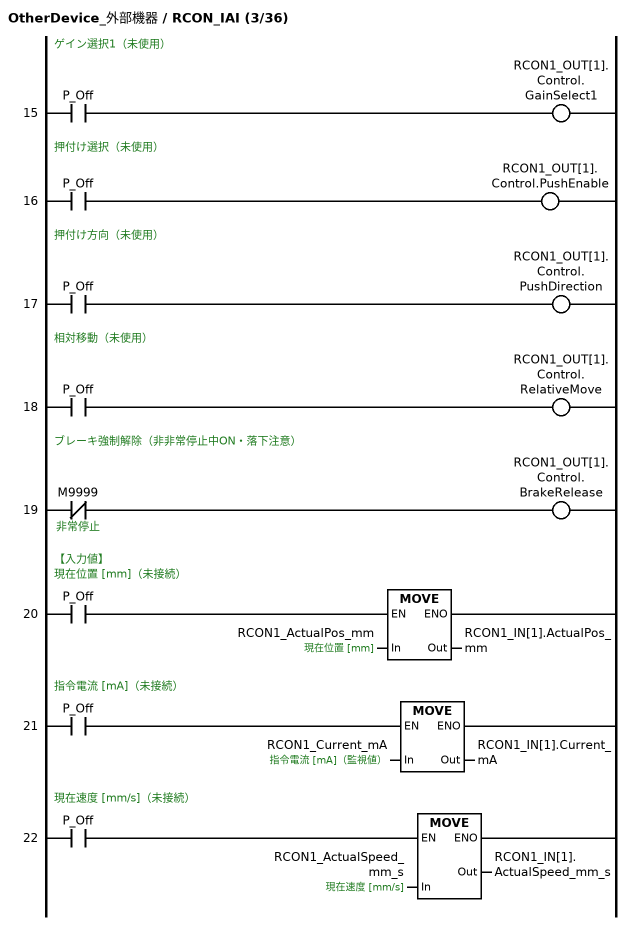
(* [picture p48: OtherDevice_外部機器 / RCON_IAI, rungs 15-22] *)
(* Rung 15: ゲイン選択1（未使用） *)
RCON1_OUT[1].Control.GainSelect1 := P_Off;
(* Rung 16: 押付け選択（未使用） *)
RCON1_OUT[1].Control.PushEnable := P_Off;
(* Rung 17: 押付け方向（未使用） *)
RCON1_OUT[1].Control.PushDirection := P_Off;
(* Rung 18: 相対移動（未使用） *)
RCON1_OUT[1].Control.RelativeMove := P_Off;
(* Rung 19: ブレーキ強制解除（非非常停止中ON・落下注意） *)
RCON1_OUT[1].Control.BrakeRelease := NOT M9999;
(* Rung 20: 【入力値】 / 現在位置 [mm]（未接続） *)
IF P_Off THEN RCON1_IN[1].ActualPos_mm := RCON1_ActualPos_mm; END_IF;
(* Rung 21: 指令電流 [mA]（未接続） *)
IF P_Off THEN RCON1_IN[1].Current_mA := RCON1_Current_mA; END_IF;
(* Rung 22: 現在速度 [mm/s]（未接続） *)
IF P_Off THEN RCON1_IN[1].ActualSpeed_mm_s := RCON1_ActualSpeed_mm_s; END_IF;

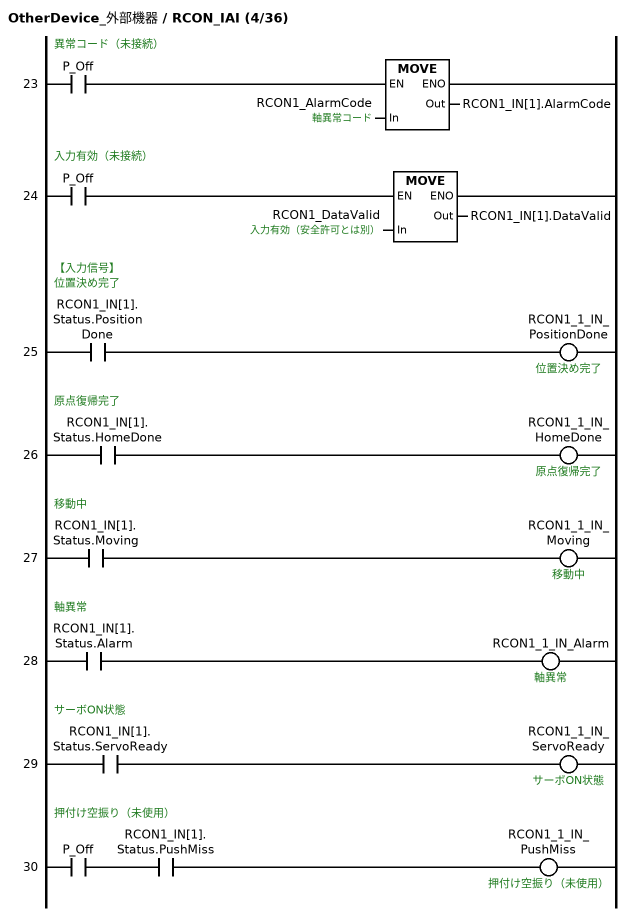
(* Rung 23: 異常コード（未接続） *)
IF P_Off THEN RCON1_IN[1].AlarmCode := RCON1_AlarmCode; END_IF;
(* Rung 24: 入力有効（未接続） *)
IF P_Off THEN RCON1_IN[1].DataValid := RCON1_DataValid; END_IF;
(* Rung 25: 【入力信号】 / 位置決め完了 *)
RCON1_1_IN_PositionDone := RCON1_IN[1].Status.PositionDone;
(* Rung 26: 原点復帰完了 *)
RCON1_1_IN_HomeDone := RCON1_IN[1].Status.HomeDone;
(* Rung 27: 移動中 *)
RCON1_1_IN_Moving := RCON1_IN[1].Status.Moving;
(* Rung 28: 軸異常 *)
RCON1_1_IN_Alarm := RCON1_IN[1].Status.Alarm;
(* Rung 29: サーボON状態 *)
RCON1_1_IN_ServoReady := RCON1_IN[1].Status.ServoReady;
(* Rung 30: 押付け空振り（未使用） *)
RCON1_1_IN_PushMiss := P_Off AND RCON1_IN[1].Status.PushMiss;

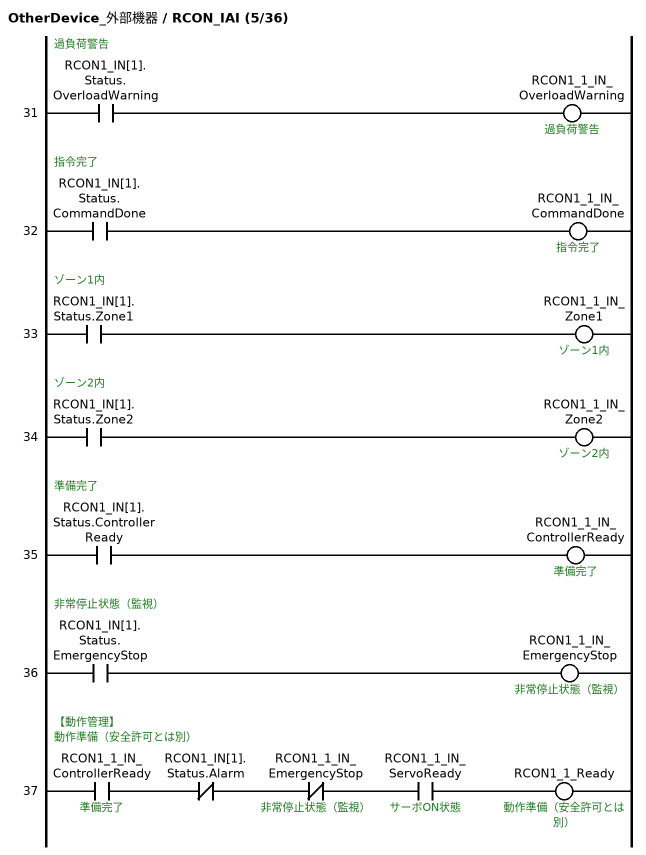
(* Rung 31: 過負荷警告 *)
RCON1_1_IN_OverloadWarning := RCON1_IN[1].Status.OverloadWarning;
(* Rung 32: 指令完了 *)
RCON1_1_IN_CommandDone := RCON1_IN[1].Status.CommandDone;
(* Rung 33: ゾーン1内 *)
RCON1_1_IN_Zone1 := RCON1_IN[1].Status.Zone1;
(* Rung 34: ゾーン2内 *)
RCON1_1_IN_Zone2 := RCON1_IN[1].Status.Zone2;
(* Rung 35: 準備完了 *)
RCON1_1_IN_ControllerReady := RCON1_IN[1].Status.ControllerReady;
(* Rung 36: 非常停止状態（監視） *)
RCON1_1_IN_EmergencyStop := RCON1_IN[1].Status.EmergencyStop;
(* Rung 37: 【動作管理】 / 動作準備（安全許可とは別） *)
RCON1_1_Ready := RCON1_1_IN_ControllerReady AND NOT RCON1_IN[1].Status.Alarm AND NOT RCON1_1_IN_EmergencyStop AND RCON1_1_IN_ServoReady;

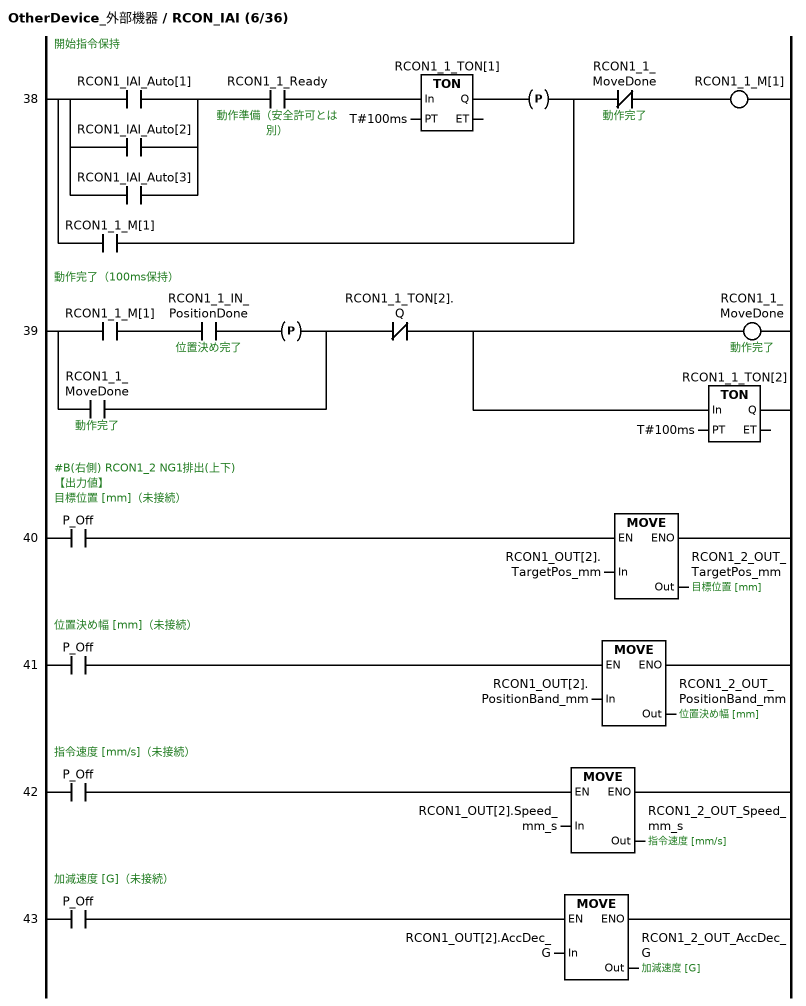
(* Rung 38: 開始指令保持 *)
RCON1_1_TON[1](In := (RCON1_IAI_Auto[1] OR RCON1_IAI_Auto[2] OR RCON1_IAI_Auto[3]) AND RCON1_1_Ready, PT := T#100ms);
_e2(CLK := RCON1_1_TON[1].Q);
RCON1_1_M[1] := (_e2.Q OR RCON1_1_M[1]) AND NOT RCON1_1_MoveDone;
(* Rung 39: 動作完了（100ms保持） *)
_e3(CLK := RCON1_1_M[1] AND RCON1_1_IN_PositionDone);
_p4 := (_e3.Q OR RCON1_1_MoveDone) AND NOT RCON1_1_TON[2].Q;
RCON1_1_MoveDone := _p4;
RCON1_1_TON[2](In := _p4, PT := T#100ms);
(* Rung 40: #B(右側) RCON1_2 NG1排出(上下) / 【出力値】 / 目標位置 [mm]（未接続） *)
IF P_Off THEN RCON1_2_OUT_TargetPos_mm := RCON1_OUT[2].TargetPos_mm; END_IF;
(* Rung 41: 位置決め幅 [mm]（未接続） *)
IF P_Off THEN RCON1_2_OUT_PositionBand_mm := RCON1_OUT[2].PositionBand_mm; END_IF;
(* Rung 42: 指令速度 [mm/s]（未接続） *)
IF P_Off THEN RCON1_2_OUT_Speed_mm_s := RCON1_OUT[2].Speed_mm_s; END_IF;
(* Rung 43: 加減速度 [G]（未接続） *)
IF P_Off THEN RCON1_2_OUT_AccDec_G := RCON1_OUT[2].AccDec_G; END_IF;

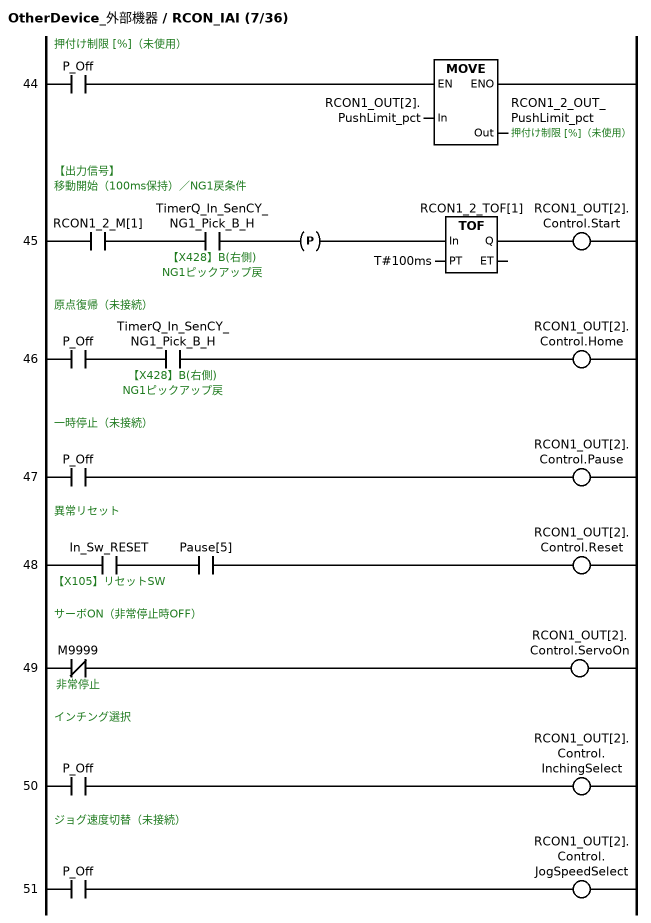
(* Rung 44: 押付け制限 [%]（未使用） *)
IF P_Off THEN RCON1_2_OUT_PushLimit_pct := RCON1_OUT[2].PushLimit_pct; END_IF;
(* Rung 45: 【出力信号】 / 移動開始（100ms保持）／NG1戻条件 *)
_e5(CLK := RCON1_2_M[1] AND TimerQ_In_SenCY_NG1_Pick_B_H);
RCON1_2_TOF[1](In := _e5.Q, PT := T#100ms);
RCON1_OUT[2].Control.Start := RCON1_2_TOF[1].Q;
(* Rung 46: 原点復帰（未接続） *)
RCON1_OUT[2].Control.Home := P_Off AND TimerQ_In_SenCY_NG1_Pick_B_H;
(* Rung 47: 一時停止（未接続） *)
RCON1_OUT[2].Control.Pause := P_Off;
(* Rung 48: 異常リセット *)
RCON1_OUT[2].Control.Reset := In_Sw_RESET AND Pause[5];
(* Rung 49: サーボON（非常停止時OFF） *)
RCON1_OUT[2].Control.ServoOn := NOT M9999;
(* Rung 50: インチング選択 *)
RCON1_OUT[2].Control.InchingSelect := P_Off;
(* Rung 51: ジョグ速度切替（未接続） *)
RCON1_OUT[2].Control.JogSpeedSelect := P_Off;

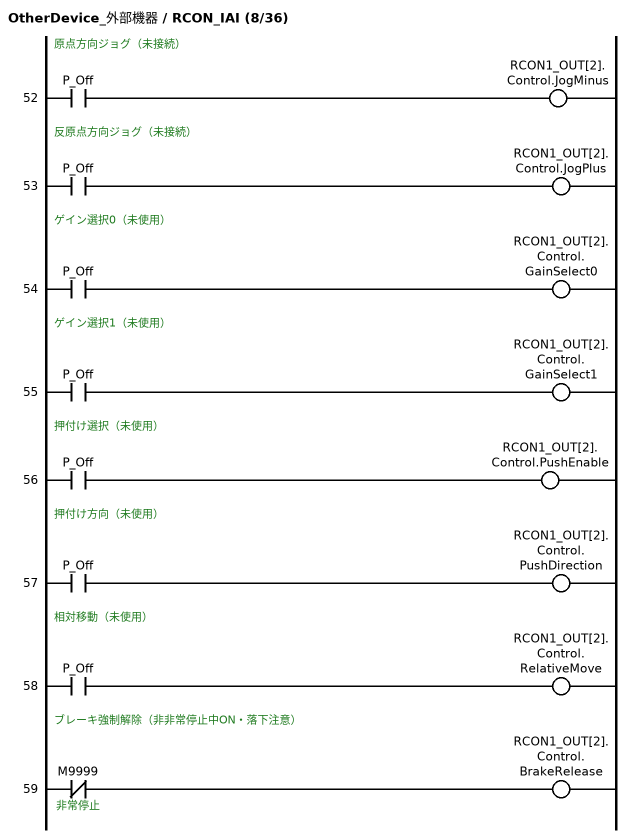
(* Rung 52: 原点方向ジョグ（未接続） *)
RCON1_OUT[2].Control.JogMinus := P_Off;
(* Rung 53: 反原点方向ジョグ（未接続） *)
RCON1_OUT[2].Control.JogPlus := P_Off;
(* Rung 54: ゲイン選択0（未使用） *)
RCON1_OUT[2].Control.GainSelect0 := P_Off;
(* Rung 55: ゲイン選択1（未使用） *)
RCON1_OUT[2].Control.GainSelect1 := P_Off;
(* Rung 56: 押付け選択（未使用） *)
RCON1_OUT[2].Control.PushEnable := P_Off;
(* Rung 57: 押付け方向（未使用） *)
RCON1_OUT[2].Control.PushDirection := P_Off;
(* Rung 58: 相対移動（未使用） *)
RCON1_OUT[2].Control.RelativeMove := P_Off;
(* Rung 59: ブレーキ強制解除（非非常停止中ON・落下注意） *)
RCON1_OUT[2].Control.BrakeRelease := NOT M9999;

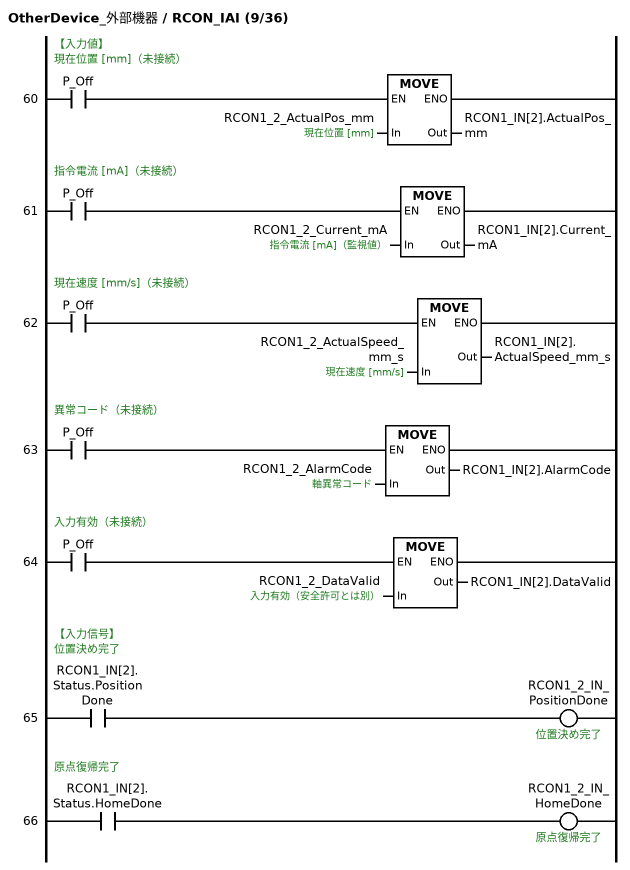
(* Rung 60: 【入力値】 / 現在位置 [mm]（未接続） *)
IF P_Off THEN RCON1_IN[2].ActualPos_mm := RCON1_2_ActualPos_mm; END_IF;
(* Rung 61: 指令電流 [mA]（未接続） *)
IF P_Off THEN RCON1_IN[2].Current_mA := RCON1_2_Current_mA; END_IF;
(* Rung 62: 現在速度 [mm/s]（未接続） *)
IF P_Off THEN RCON1_IN[2].ActualSpeed_mm_s := RCON1_2_ActualSpeed_mm_s; END_IF;
(* Rung 63: 異常コード（未接続） *)
IF P_Off THEN RCON1_IN[2].AlarmCode := RCON1_2_AlarmCode; END_IF;
(* Rung 64: 入力有効（未接続） *)
IF P_Off THEN RCON1_IN[2].DataValid := RCON1_2_DataValid; END_IF;
(* Rung 65: 【入力信号】 / 位置決め完了 *)
RCON1_2_IN_PositionDone := RCON1_IN[2].Status.PositionDone;
(* Rung 66: 原点復帰完了 *)
RCON1_2_IN_HomeDone := RCON1_IN[2].Status.HomeDone;

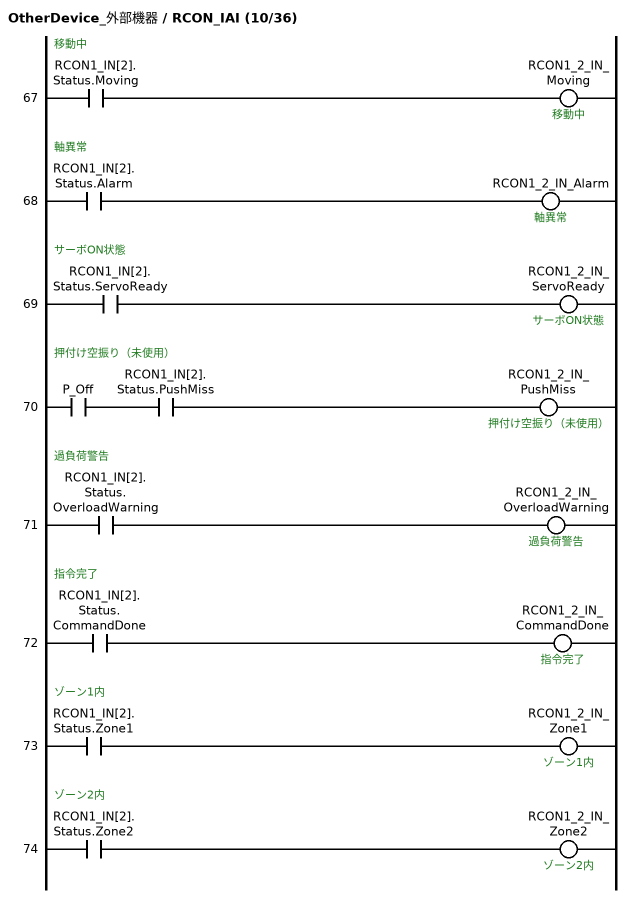
(* Rung 67: 移動中 *)
RCON1_2_IN_Moving := RCON1_IN[2].Status.Moving;
(* Rung 68: 軸異常 *)
RCON1_2_IN_Alarm := RCON1_IN[2].Status.Alarm;
(* Rung 69: サーボON状態 *)
RCON1_2_IN_ServoReady := RCON1_IN[2].Status.ServoReady;
(* Rung 70: 押付け空振り（未使用） *)
RCON1_2_IN_PushMiss := P_Off AND RCON1_IN[2].Status.PushMiss;
(* Rung 71: 過負荷警告 *)
RCON1_2_IN_OverloadWarning := RCON1_IN[2].Status.OverloadWarning;
(* Rung 72: 指令完了 *)
RCON1_2_IN_CommandDone := RCON1_IN[2].Status.CommandDone;
(* Rung 73: ゾーン1内 *)
RCON1_2_IN_Zone1 := RCON1_IN[2].Status.Zone1;
(* Rung 74: ゾーン2内 *)
RCON1_2_IN_Zone2 := RCON1_IN[2].Status.Zone2;

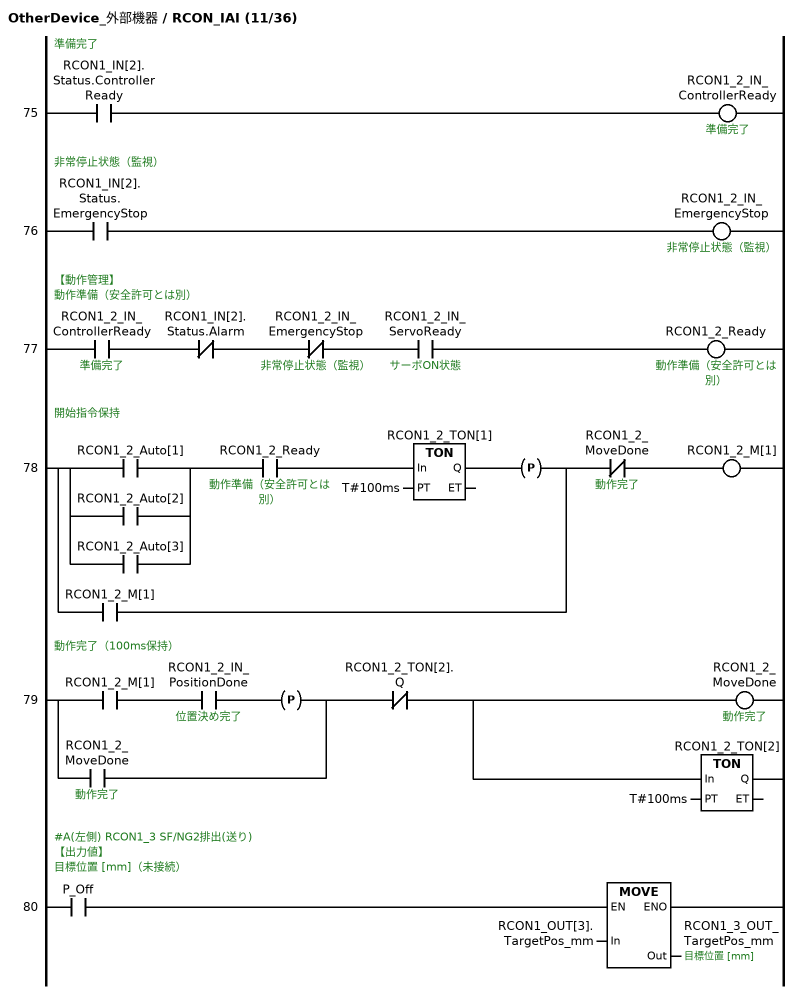
(* Rung 75: 準備完了 *)
RCON1_2_IN_ControllerReady := RCON1_IN[2].Status.ControllerReady;
(* Rung 76: 非常停止状態（監視） *)
RCON1_2_IN_EmergencyStop := RCON1_IN[2].Status.EmergencyStop;
(* Rung 77: 【動作管理】 / 動作準備（安全許可とは別） *)
RCON1_2_Ready := RCON1_2_IN_ControllerReady AND NOT RCON1_IN[2].Status.Alarm AND NOT RCON1_2_IN_EmergencyStop AND RCON1_2_IN_ServoReady;
(* Rung 78: 開始指令保持 *)
RCON1_2_TON[1](In := (RCON1_2_Auto[1] OR RCON1_2_Auto[2] OR RCON1_2_Auto[3]) AND RCON1_2_Ready, PT := T#100ms);
_e6(CLK := RCON1_2_TON[1].Q);
RCON1_2_M[1] := (_e6.Q OR RCON1_2_M[1]) AND NOT RCON1_2_MoveDone;
(* Rung 79: 動作完了（100ms保持） *)
_e7(CLK := RCON1_2_M[1] AND RCON1_2_IN_PositionDone);
_p8 := (_e7.Q OR RCON1_2_MoveDone) AND NOT RCON1_2_TON[2].Q;
RCON1_2_MoveDone := _p8;
RCON1_2_TON[2](In := _p8, PT := T#100ms);
(* Rung 80: #A(左側) RCON1_3 SF/NG2排出(送り) / 【出力値】 / 目標位置 [mm]（未接続） *)
IF P_Off THEN RCON1_3_OUT_TargetPos_mm := RCON1_OUT[3].TargetPos_mm; END_IF;

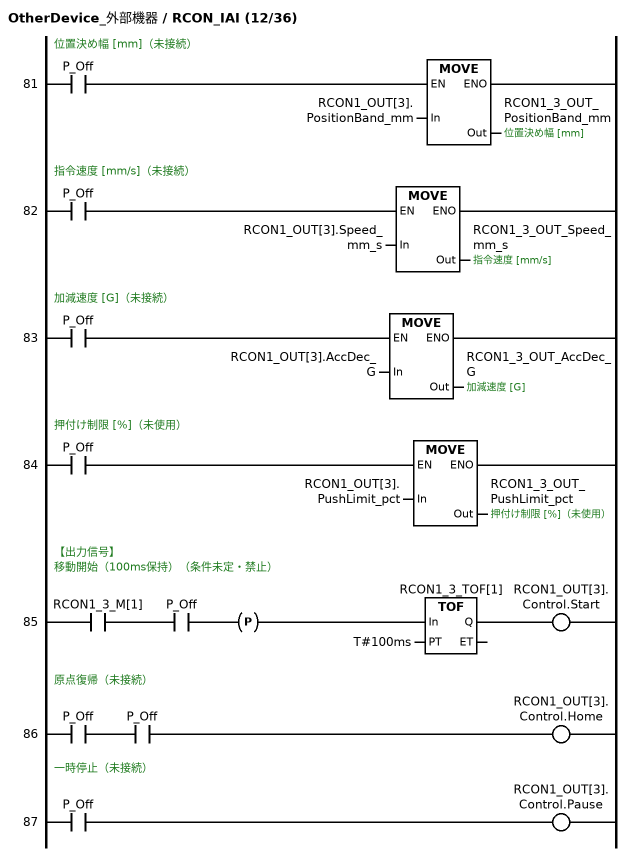
(* Rung 81: 位置決め幅 [mm]（未接続） *)
IF P_Off THEN RCON1_3_OUT_PositionBand_mm := RCON1_OUT[3].PositionBand_mm; END_IF;
(* Rung 82: 指令速度 [mm/s]（未接続） *)
IF P_Off THEN RCON1_3_OUT_Speed_mm_s := RCON1_OUT[3].Speed_mm_s; END_IF;
(* Rung 83: 加減速度 [G]（未接続） *)
IF P_Off THEN RCON1_3_OUT_AccDec_G := RCON1_OUT[3].AccDec_G; END_IF;
(* Rung 84: 押付け制限 [%]（未使用） *)
IF P_Off THEN RCON1_3_OUT_PushLimit_pct := RCON1_OUT[3].PushLimit_pct; END_IF;
(* Rung 85: 【出力信号】 / 移動開始（100ms保持）（条件未定・禁止） *)
_e9(CLK := RCON1_3_M[1] AND P_Off);
RCON1_3_TOF[1](In := _e9.Q, PT := T#100ms);
RCON1_OUT[3].Control.Start := RCON1_3_TOF[1].Q;
(* Rung 86: 原点復帰（未接続） *)
RCON1_OUT[3].Control.Home := P_Off AND P_Off;
(* Rung 87: 一時停止（未接続） *)
RCON1_OUT[3].Control.Pause := P_Off;

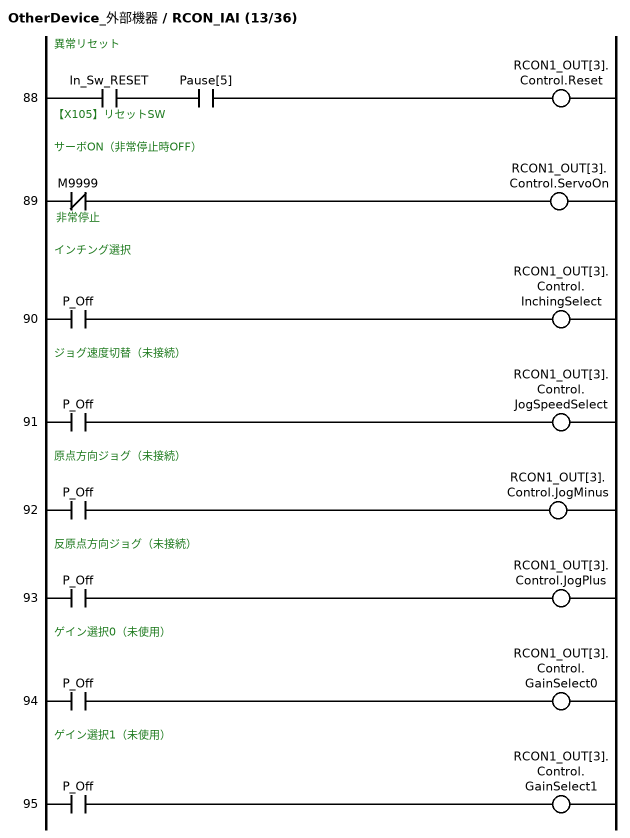
(* Rung 88: 異常リセット *)
RCON1_OUT[3].Control.Reset := In_Sw_RESET AND Pause[5];
(* Rung 89: サーボON（非常停止時OFF） *)
RCON1_OUT[3].Control.ServoOn := NOT M9999;
(* Rung 90: インチング選択 *)
RCON1_OUT[3].Control.InchingSelect := P_Off;
(* Rung 91: ジョグ速度切替（未接続） *)
RCON1_OUT[3].Control.JogSpeedSelect := P_Off;
(* Rung 92: 原点方向ジョグ（未接続） *)
RCON1_OUT[3].Control.JogMinus := P_Off;
(* Rung 93: 反原点方向ジョグ（未接続） *)
RCON1_OUT[3].Control.JogPlus := P_Off;
(* Rung 94: ゲイン選択0（未使用） *)
RCON1_OUT[3].Control.GainSelect0 := P_Off;
(* Rung 95: ゲイン選択1（未使用） *)
RCON1_OUT[3].Control.GainSelect1 := P_Off;

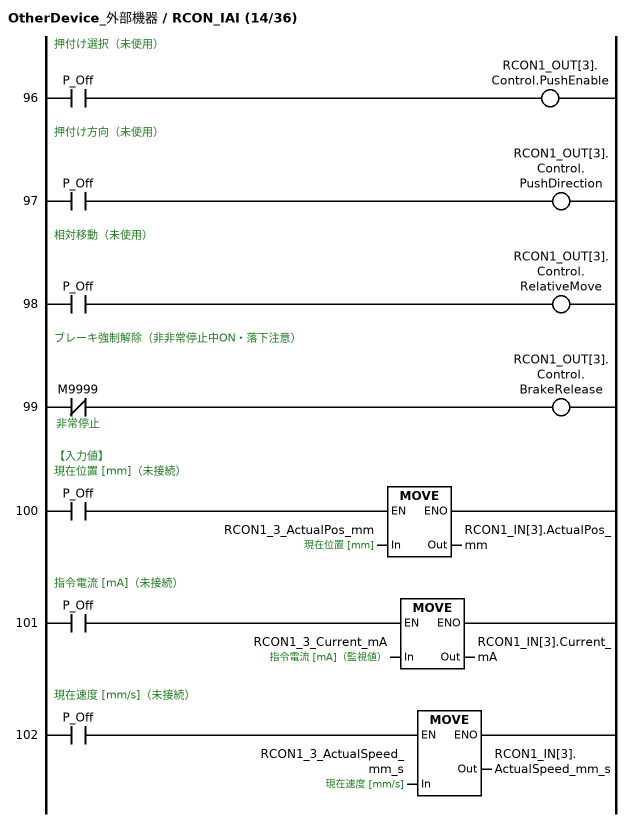
(* Rung 96: 押付け選択（未使用） *)
RCON1_OUT[3].Control.PushEnable := P_Off;
(* Rung 97: 押付け方向（未使用） *)
RCON1_OUT[3].Control.PushDirection := P_Off;
(* Rung 98: 相対移動（未使用） *)
RCON1_OUT[3].Control.RelativeMove := P_Off;
(* Rung 99: ブレーキ強制解除（非非常停止中ON・落下注意） *)
RCON1_OUT[3].Control.BrakeRelease := NOT M9999;
(* Rung 100: 【入力値】 / 現在位置 [mm]（未接続） *)
IF P_Off THEN RCON1_IN[3].ActualPos_mm := RCON1_3_ActualPos_mm; END_IF;
(* Rung 101: 指令電流 [mA]（未接続） *)
IF P_Off THEN RCON1_IN[3].Current_mA := RCON1_3_Current_mA; END_IF;
(* Rung 102: 現在速度 [mm/s]（未接続） *)
IF P_Off THEN RCON1_IN[3].ActualSpeed_mm_s := RCON1_3_ActualSpeed_mm_s; END_IF;

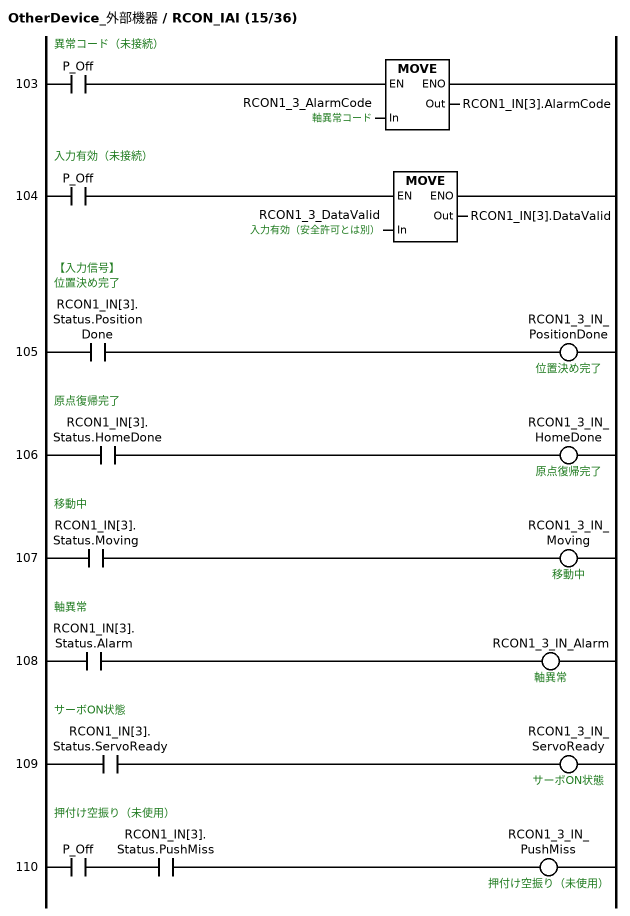
(* Rung 103: 異常コード（未接続） *)
IF P_Off THEN RCON1_IN[3].AlarmCode := RCON1_3_AlarmCode; END_IF;
(* Rung 104: 入力有効（未接続） *)
IF P_Off THEN RCON1_IN[3].DataValid := RCON1_3_DataValid; END_IF;
(* Rung 105: 【入力信号】 / 位置決め完了 *)
RCON1_3_IN_PositionDone := RCON1_IN[3].Status.PositionDone;
(* Rung 106: 原点復帰完了 *)
RCON1_3_IN_HomeDone := RCON1_IN[3].Status.HomeDone;
(* Rung 107: 移動中 *)
RCON1_3_IN_Moving := RCON1_IN[3].Status.Moving;
(* Rung 108: 軸異常 *)
RCON1_3_IN_Alarm := RCON1_IN[3].Status.Alarm;
(* Rung 109: サーボON状態 *)
RCON1_3_IN_ServoReady := RCON1_IN[3].Status.ServoReady;
(* Rung 110: 押付け空振り（未使用） *)
RCON1_3_IN_PushMiss := P_Off AND RCON1_IN[3].Status.PushMiss;

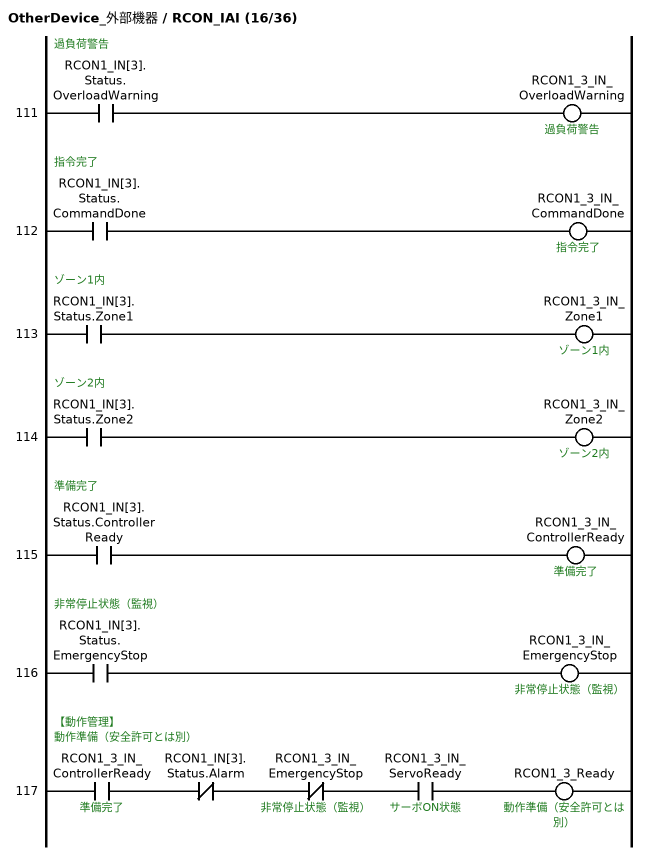
(* Rung 111: 過負荷警告 *)
RCON1_3_IN_OverloadWarning := RCON1_IN[3].Status.OverloadWarning;
(* Rung 112: 指令完了 *)
RCON1_3_IN_CommandDone := RCON1_IN[3].Status.CommandDone;
(* Rung 113: ゾーン1内 *)
RCON1_3_IN_Zone1 := RCON1_IN[3].Status.Zone1;
(* Rung 114: ゾーン2内 *)
RCON1_3_IN_Zone2 := RCON1_IN[3].Status.Zone2;
(* Rung 115: 準備完了 *)
RCON1_3_IN_ControllerReady := RCON1_IN[3].Status.ControllerReady;
(* Rung 116: 非常停止状態（監視） *)
RCON1_3_IN_EmergencyStop := RCON1_IN[3].Status.EmergencyStop;
(* Rung 117: 【動作管理】 / 動作準備（安全許可とは別） *)
RCON1_3_Ready := RCON1_3_IN_ControllerReady AND NOT RCON1_IN[3].Status.Alarm AND NOT RCON1_3_IN_EmergencyStop AND RCON1_3_IN_ServoReady;

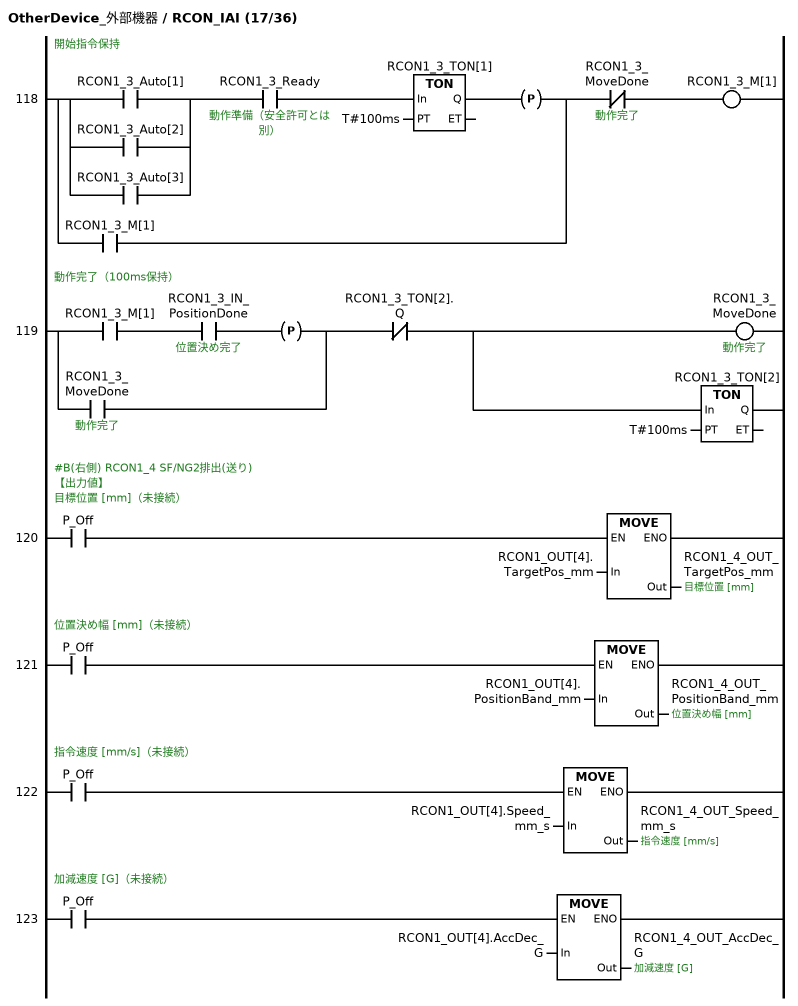
(* Rung 118: 開始指令保持 *)
RCON1_3_TON[1](In := (RCON1_3_Auto[1] OR RCON1_3_Auto[2] OR RCON1_3_Auto[3]) AND RCON1_3_Ready, PT := T#100ms);
_e10(CLK := RCON1_3_TON[1].Q);
RCON1_3_M[1] := (_e10.Q OR RCON1_3_M[1]) AND NOT RCON1_3_MoveDone;
(* Rung 119: 動作完了（100ms保持） *)
_e11(CLK := RCON1_3_M[1] AND RCON1_3_IN_PositionDone);
_p12 := (_e11.Q OR RCON1_3_MoveDone) AND NOT RCON1_3_TON[2].Q;
RCON1_3_MoveDone := _p12;
RCON1_3_TON[2](In := _p12, PT := T#100ms);
(* Rung 120: #B(右側) RCON1_4 SF/NG2排出(送り) / 【出力値】 / 目標位置 [mm]（未接続） *)
IF P_Off THEN RCON1_4_OUT_TargetPos_mm := RCON1_OUT[4].TargetPos_mm; END_IF;
(* Rung 121: 位置決め幅 [mm]（未接続） *)
IF P_Off THEN RCON1_4_OUT_PositionBand_mm := RCON1_OUT[4].PositionBand_mm; END_IF;
(* Rung 122: 指令速度 [mm/s]（未接続） *)
IF P_Off THEN RCON1_4_OUT_Speed_mm_s := RCON1_OUT[4].Speed_mm_s; END_IF;
(* Rung 123: 加減速度 [G]（未接続） *)
IF P_Off THEN RCON1_4_OUT_AccDec_G := RCON1_OUT[4].AccDec_G; END_IF;

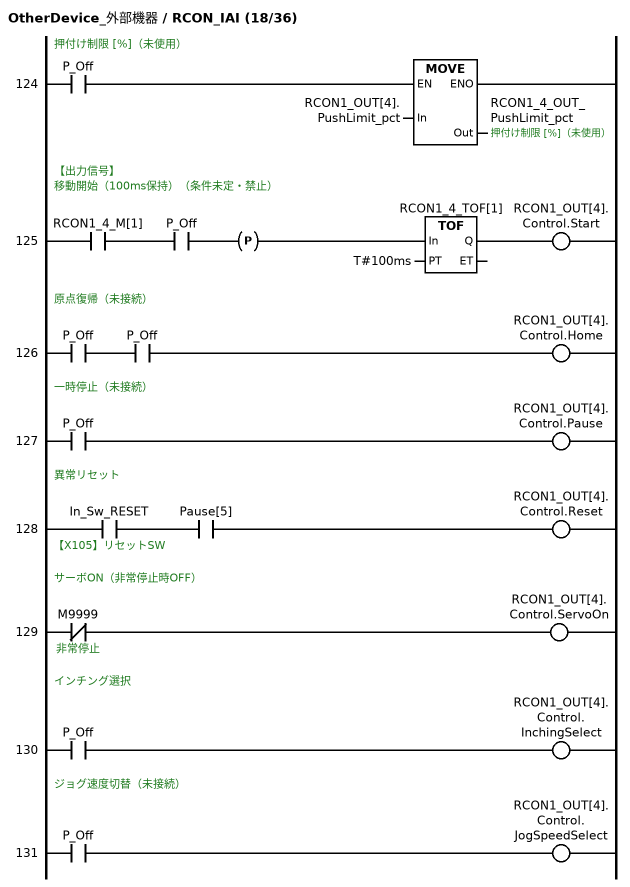
(* Rung 124: 押付け制限 [%]（未使用） *)
IF P_Off THEN RCON1_4_OUT_PushLimit_pct := RCON1_OUT[4].PushLimit_pct; END_IF;
(* Rung 125: 【出力信号】 / 移動開始（100ms保持）（条件未定・禁止） *)
_e13(CLK := RCON1_4_M[1] AND P_Off);
RCON1_4_TOF[1](In := _e13.Q, PT := T#100ms);
RCON1_OUT[4].Control.Start := RCON1_4_TOF[1].Q;
(* Rung 126: 原点復帰（未接続） *)
RCON1_OUT[4].Control.Home := P_Off AND P_Off;
(* Rung 127: 一時停止（未接続） *)
RCON1_OUT[4].Control.Pause := P_Off;
(* Rung 128: 異常リセット *)
RCON1_OUT[4].Control.Reset := In_Sw_RESET AND Pause[5];
(* Rung 129: サーボON（非常停止時OFF） *)
RCON1_OUT[4].Control.ServoOn := NOT M9999;
(* Rung 130: インチング選択 *)
RCON1_OUT[4].Control.InchingSelect := P_Off;
(* Rung 131: ジョグ速度切替（未接続） *)
RCON1_OUT[4].Control.JogSpeedSelect := P_Off;

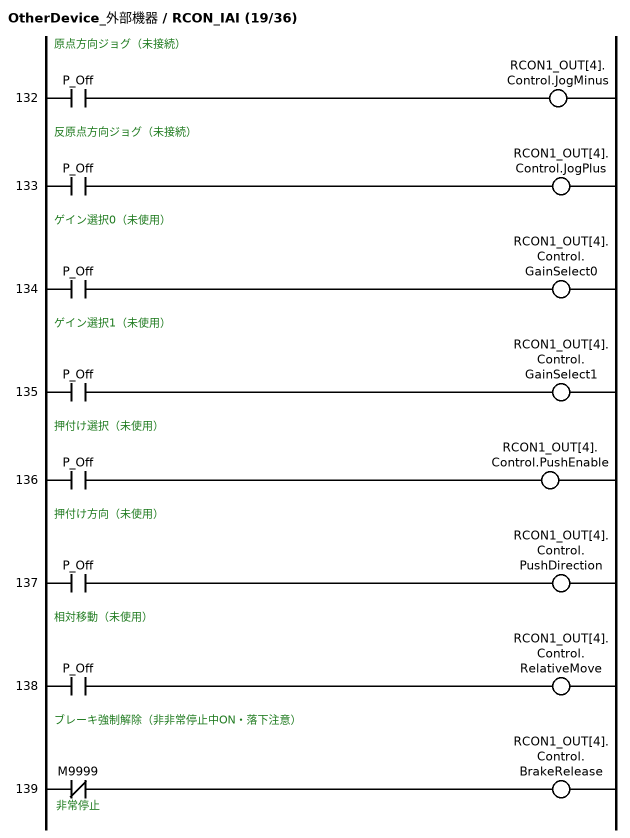
(* Rung 132: 原点方向ジョグ（未接続） *)
RCON1_OUT[4].Control.JogMinus := P_Off;
(* Rung 133: 反原点方向ジョグ（未接続） *)
RCON1_OUT[4].Control.JogPlus := P_Off;
(* Rung 134: ゲイン選択0（未使用） *)
RCON1_OUT[4].Control.GainSelect0 := P_Off;
(* Rung 135: ゲイン選択1（未使用） *)
RCON1_OUT[4].Control.GainSelect1 := P_Off;
(* Rung 136: 押付け選択（未使用） *)
RCON1_OUT[4].Control.PushEnable := P_Off;
(* Rung 137: 押付け方向（未使用） *)
RCON1_OUT[4].Control.PushDirection := P_Off;
(* Rung 138: 相対移動（未使用） *)
RCON1_OUT[4].Control.RelativeMove := P_Off;
(* Rung 139: ブレーキ強制解除（非非常停止中ON・落下注意） *)
RCON1_OUT[4].Control.BrakeRelease := NOT M9999;

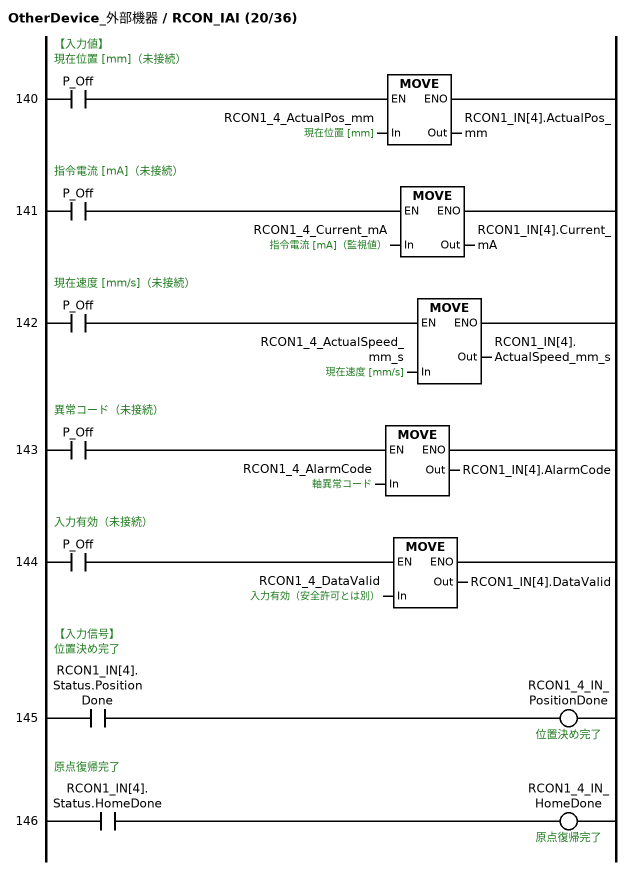
(* Rung 140: 【入力値】 / 現在位置 [mm]（未接続） *)
IF P_Off THEN RCON1_IN[4].ActualPos_mm := RCON1_4_ActualPos_mm; END_IF;
(* Rung 141: 指令電流 [mA]（未接続） *)
IF P_Off THEN RCON1_IN[4].Current_mA := RCON1_4_Current_mA; END_IF;
(* Rung 142: 現在速度 [mm/s]（未接続） *)
IF P_Off THEN RCON1_IN[4].ActualSpeed_mm_s := RCON1_4_ActualSpeed_mm_s; END_IF;
(* Rung 143: 異常コード（未接続） *)
IF P_Off THEN RCON1_IN[4].AlarmCode := RCON1_4_AlarmCode; END_IF;
(* Rung 144: 入力有効（未接続） *)
IF P_Off THEN RCON1_IN[4].DataValid := RCON1_4_DataValid; END_IF;
(* Rung 145: 【入力信号】 / 位置決め完了 *)
RCON1_4_IN_PositionDone := RCON1_IN[4].Status.PositionDone;
(* Rung 146: 原点復帰完了 *)
RCON1_4_IN_HomeDone := RCON1_IN[4].Status.HomeDone;

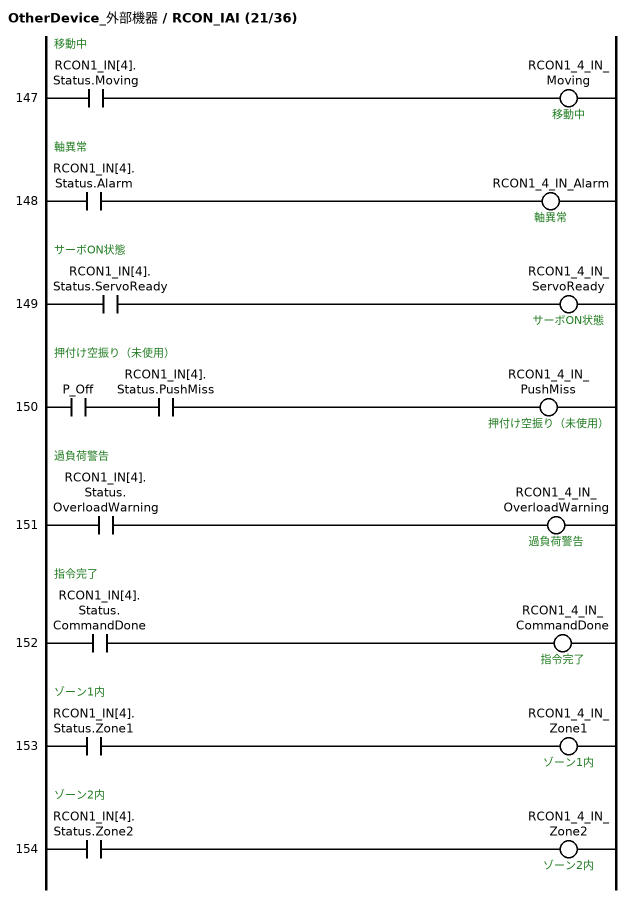
(* Rung 147: 移動中 *)
RCON1_4_IN_Moving := RCON1_IN[4].Status.Moving;
(* Rung 148: 軸異常 *)
RCON1_4_IN_Alarm := RCON1_IN[4].Status.Alarm;
(* Rung 149: サーボON状態 *)
RCON1_4_IN_ServoReady := RCON1_IN[4].Status.ServoReady;
(* Rung 150: 押付け空振り（未使用） *)
RCON1_4_IN_PushMiss := P_Off AND RCON1_IN[4].Status.PushMiss;
(* Rung 151: 過負荷警告 *)
RCON1_4_IN_OverloadWarning := RCON1_IN[4].Status.OverloadWarning;
(* Rung 152: 指令完了 *)
RCON1_4_IN_CommandDone := RCON1_IN[4].Status.CommandDone;
(* Rung 153: ゾーン1内 *)
RCON1_4_IN_Zone1 := RCON1_IN[4].Status.Zone1;
(* Rung 154: ゾーン2内 *)
RCON1_4_IN_Zone2 := RCON1_IN[4].Status.Zone2;

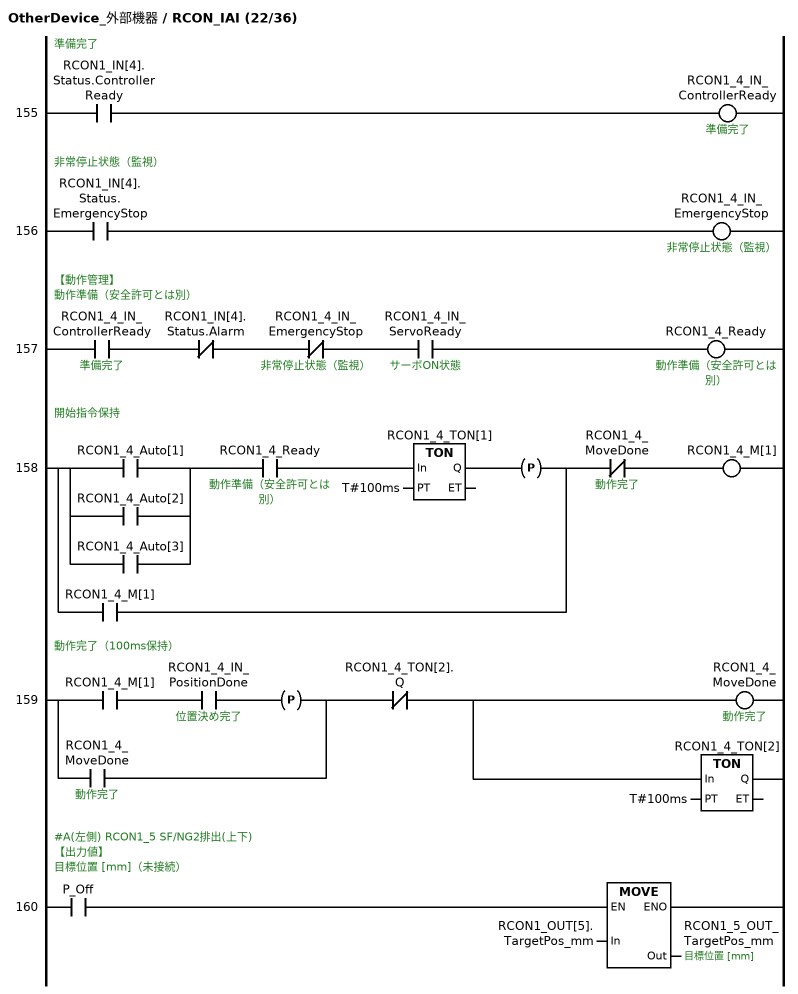
(* Rung 155: 準備完了 *)
RCON1_4_IN_ControllerReady := RCON1_IN[4].Status.ControllerReady;
(* Rung 156: 非常停止状態（監視） *)
RCON1_4_IN_EmergencyStop := RCON1_IN[4].Status.EmergencyStop;
(* Rung 157: 【動作管理】 / 動作準備（安全許可とは別） *)
RCON1_4_Ready := RCON1_4_IN_ControllerReady AND NOT RCON1_IN[4].Status.Alarm AND NOT RCON1_4_IN_EmergencyStop AND RCON1_4_IN_ServoReady;
(* Rung 158: 開始指令保持 *)
RCON1_4_TON[1](In := (RCON1_4_Auto[1] OR RCON1_4_Auto[2] OR RCON1_4_Auto[3]) AND RCON1_4_Ready, PT := T#100ms);
_e14(CLK := RCON1_4_TON[1].Q);
RCON1_4_M[1] := (_e14.Q OR RCON1_4_M[1]) AND NOT RCON1_4_MoveDone;
(* Rung 159: 動作完了（100ms保持） *)
_e15(CLK := RCON1_4_M[1] AND RCON1_4_IN_PositionDone);
_p16 := (_e15.Q OR RCON1_4_MoveDone) AND NOT RCON1_4_TON[2].Q;
RCON1_4_MoveDone := _p16;
RCON1_4_TON[2](In := _p16, PT := T#100ms);
(* Rung 160: #A(左側) RCON1_5 SF/NG2排出(上下) / 【出力値】 / 目標位置 [mm]（未接続） *)
IF P_Off THEN RCON1_5_OUT_TargetPos_mm := RCON1_OUT[5].TargetPos_mm; END_IF;

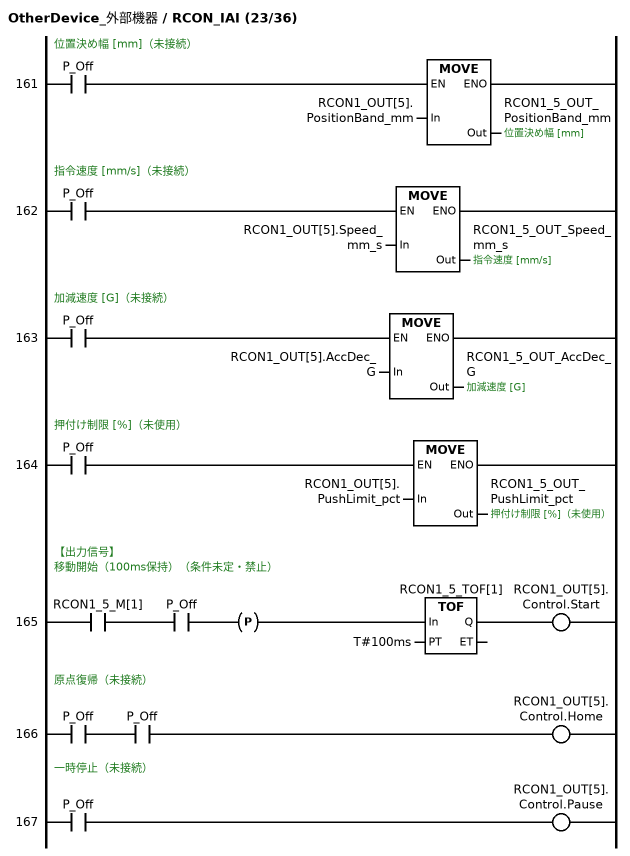
(* Rung 161: 位置決め幅 [mm]（未接続） *)
IF P_Off THEN RCON1_5_OUT_PositionBand_mm := RCON1_OUT[5].PositionBand_mm; END_IF;
(* Rung 162: 指令速度 [mm/s]（未接続） *)
IF P_Off THEN RCON1_5_OUT_Speed_mm_s := RCON1_OUT[5].Speed_mm_s; END_IF;
(* Rung 163: 加減速度 [G]（未接続） *)
IF P_Off THEN RCON1_5_OUT_AccDec_G := RCON1_OUT[5].AccDec_G; END_IF;
(* Rung 164: 押付け制限 [%]（未使用） *)
IF P_Off THEN RCON1_5_OUT_PushLimit_pct := RCON1_OUT[5].PushLimit_pct; END_IF;
(* Rung 165: 【出力信号】 / 移動開始（100ms保持）（条件未定・禁止） *)
_e17(CLK := RCON1_5_M[1] AND P_Off);
RCON1_5_TOF[1](In := _e17.Q, PT := T#100ms);
RCON1_OUT[5].Control.Start := RCON1_5_TOF[1].Q;
(* Rung 166: 原点復帰（未接続） *)
RCON1_OUT[5].Control.Home := P_Off AND P_Off;
(* Rung 167: 一時停止（未接続） *)
RCON1_OUT[5].Control.Pause := P_Off;

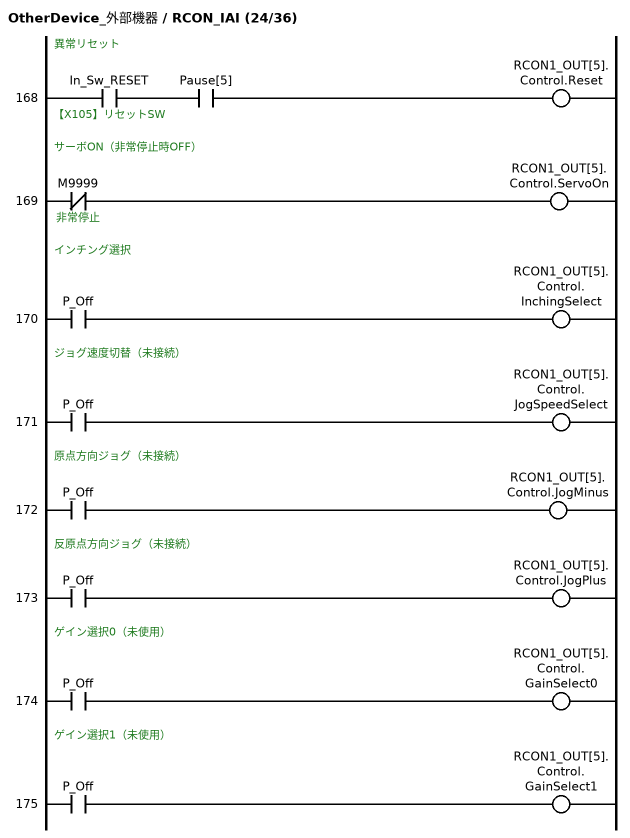
(* Rung 168: 異常リセット *)
RCON1_OUT[5].Control.Reset := In_Sw_RESET AND Pause[5];
(* Rung 169: サーボON（非常停止時OFF） *)
RCON1_OUT[5].Control.ServoOn := NOT M9999;
(* Rung 170: インチング選択 *)
RCON1_OUT[5].Control.InchingSelect := P_Off;
(* Rung 171: ジョグ速度切替（未接続） *)
RCON1_OUT[5].Control.JogSpeedSelect := P_Off;
(* Rung 172: 原点方向ジョグ（未接続） *)
RCON1_OUT[5].Control.JogMinus := P_Off;
(* Rung 173: 反原点方向ジョグ（未接続） *)
RCON1_OUT[5].Control.JogPlus := P_Off;
(* Rung 174: ゲイン選択0（未使用） *)
RCON1_OUT[5].Control.GainSelect0 := P_Off;
(* Rung 175: ゲイン選択1（未使用） *)
RCON1_OUT[5].Control.GainSelect1 := P_Off;

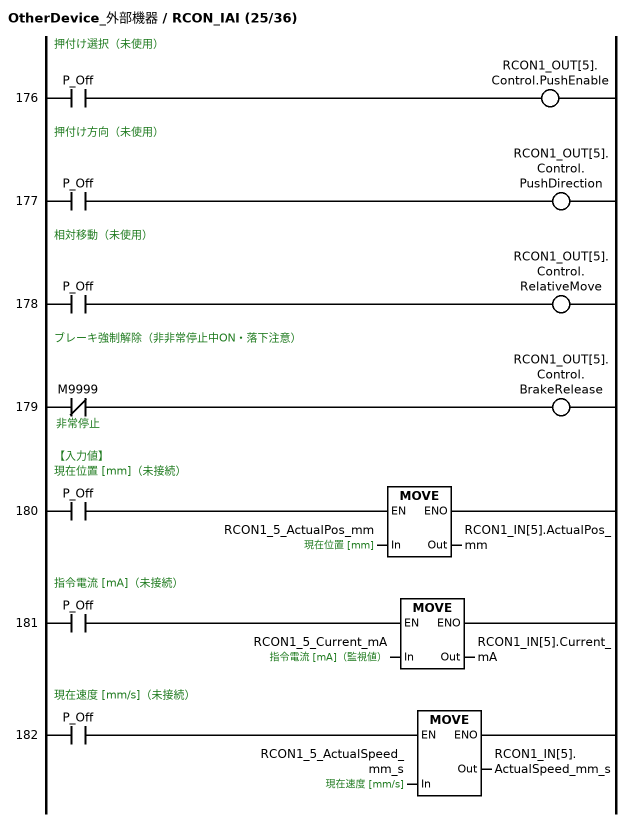
(* Rung 176: 押付け選択（未使用） *)
RCON1_OUT[5].Control.PushEnable := P_Off;
(* Rung 177: 押付け方向（未使用） *)
RCON1_OUT[5].Control.PushDirection := P_Off;
(* Rung 178: 相対移動（未使用） *)
RCON1_OUT[5].Control.RelativeMove := P_Off;
(* Rung 179: ブレーキ強制解除（非非常停止中ON・落下注意） *)
RCON1_OUT[5].Control.BrakeRelease := NOT M9999;
(* Rung 180: 【入力値】 / 現在位置 [mm]（未接続） *)
IF P_Off THEN RCON1_IN[5].ActualPos_mm := RCON1_5_ActualPos_mm; END_IF;
(* Rung 181: 指令電流 [mA]（未接続） *)
IF P_Off THEN RCON1_IN[5].Current_mA := RCON1_5_Current_mA; END_IF;
(* Rung 182: 現在速度 [mm/s]（未接続） *)
IF P_Off THEN RCON1_IN[5].ActualSpeed_mm_s := RCON1_5_ActualSpeed_mm_s; END_IF;

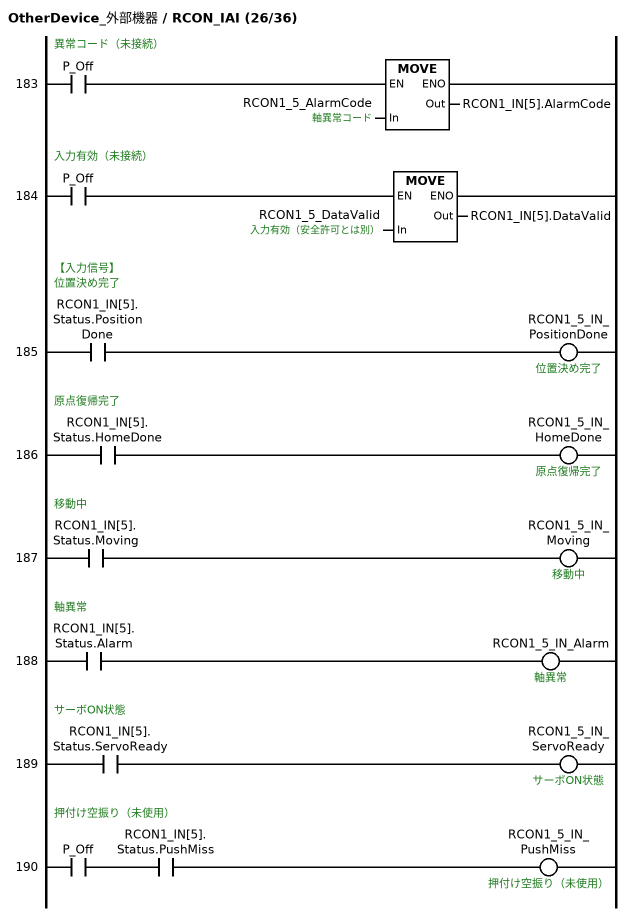
(* Rung 183: 異常コード（未接続） *)
IF P_Off THEN RCON1_IN[5].AlarmCode := RCON1_5_AlarmCode; END_IF;
(* Rung 184: 入力有効（未接続） *)
IF P_Off THEN RCON1_IN[5].DataValid := RCON1_5_DataValid; END_IF;
(* Rung 185: 【入力信号】 / 位置決め完了 *)
RCON1_5_IN_PositionDone := RCON1_IN[5].Status.PositionDone;
(* Rung 186: 原点復帰完了 *)
RCON1_5_IN_HomeDone := RCON1_IN[5].Status.HomeDone;
(* Rung 187: 移動中 *)
RCON1_5_IN_Moving := RCON1_IN[5].Status.Moving;
(* Rung 188: 軸異常 *)
RCON1_5_IN_Alarm := RCON1_IN[5].Status.Alarm;
(* Rung 189: サーボON状態 *)
RCON1_5_IN_ServoReady := RCON1_IN[5].Status.ServoReady;
(* Rung 190: 押付け空振り（未使用） *)
RCON1_5_IN_PushMiss := P_Off AND RCON1_IN[5].Status.PushMiss;

